// TIA Portal V21 export
// export: Created 2026-11-11T00:47:46.8974288Z, ExportSetting WithDefaults, DisplayName Totally Integrated Automation Portal, DisplayVersion V21 Update 3, DisplayName STEP 7 Professional, DisplayVersion V21 Update 3, DisplayName STEP 7 Safety, DisplayVersion V21, DisplayName Tech WebApplication, DisplayVersion V21, DisplayName WinCC Basic/Comfort/Advanced, DisplayVersion V21 Update 3, DisplayName WinCC Unified, DisplayVersion V21 Update 3
FUNCTION_BLOCK "FB_Fbd_sc003"   // FB182, FBD
{ S7_Optimized_Access := 'TRUE' }
VERSION : 0.1
// stored: AutoNumber true, IsIECCheckEnabled false, IsRetainMemResEnabled false, MemoryReserve 100, SetENOAutomatically false, UDAEnableTagReadback false
   VAR_INPUT
      v_req : Bool;
      v_id : CONN_PRG;
      v_r_id : CONN_R_ID;
   END_VAR
   VAR_OUTPUT
      v_done : Bool;
      v_error : Bool;
      v_status : Word;
   END_VAR
   VAR_IN_OUT
      v_sd_1 : Variant;
      v_sd_2 : Variant;
      v_sd_3 : Variant;
      v_sd_4 : Variant;
   END_VAR
   VAR
      inst { S7_SetPoint := 'True'} : USEND;
   END_VAR
BEGIN

REGION Network 1: USEND - Send data uncoordinated
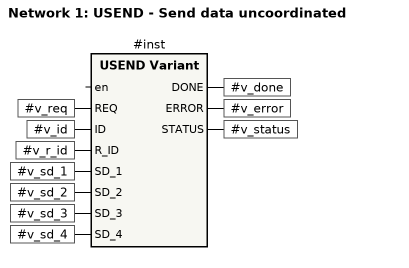
   #inst(REQ := #v_req,   // USEND
         ID := #v_id,
         R_ID := #v_r_id,
         SD_1 := #v_sd_1,
         SD_2 := #v_sd_2,
         SD_3 := #v_sd_3,
         SD_4 := #v_sd_4,
         DONE => #v_done,
         ERROR => #v_error,
         STATUS => #v_status);
END_REGION
END_FUNCTION_BLOCK
